Staubli VAL3: insertDelay.pgx

public program insertDelay(string x_sKey, num x_nIndex, bool& x_bToSave, num x_nMoveType, num x_nDelay)
  local num l_j
  local num l_i
begin
  //insert(trajTemp:tTrajItem[x_sKey].pPointItem[x_nIndex+1])
  append(trajTemp:tTrajItem[x_sKey].pPointItem)

  for l_i = (size(trajTemp:tTrajItem[x_sKey].pPointItem)-1) to(x_nIndex+1) step -1
   // logMsg(toString("",l_i))
    call copyPoint3(x_sKey,l_i,l_i-1)
  endFor
  trajTemp:tTrajItem[x_sKey].pPointItem[x_nIndex+1].pParaItem.nMoveType=x_nMoveType

  trajTemp:tTrajItem[x_sKey].pPointItem[x_nIndex+1].pParaItem.nDelay=x_nDelay

 //trajTemp:libSave()

  x_bToSave=true
end
